// TIA Portal V20 export
DATA_BLOCK "DB002_LabView_DB"   // DB3
// stored: InstanceOfName FB002_LabView, InstanceOfType FB
"FB002_LabView"
BEGIN
END_DATA_BLOCK
